Staubli VAL3: utAppearance.dtx

public string sBackgroundColour
public string sColour
public bool bVisibility
